// Mitsubishi GX Works2 project: TRANG TRAI BAN CU   PLC: FX3U/FX3UC

PROGRAM MAIN
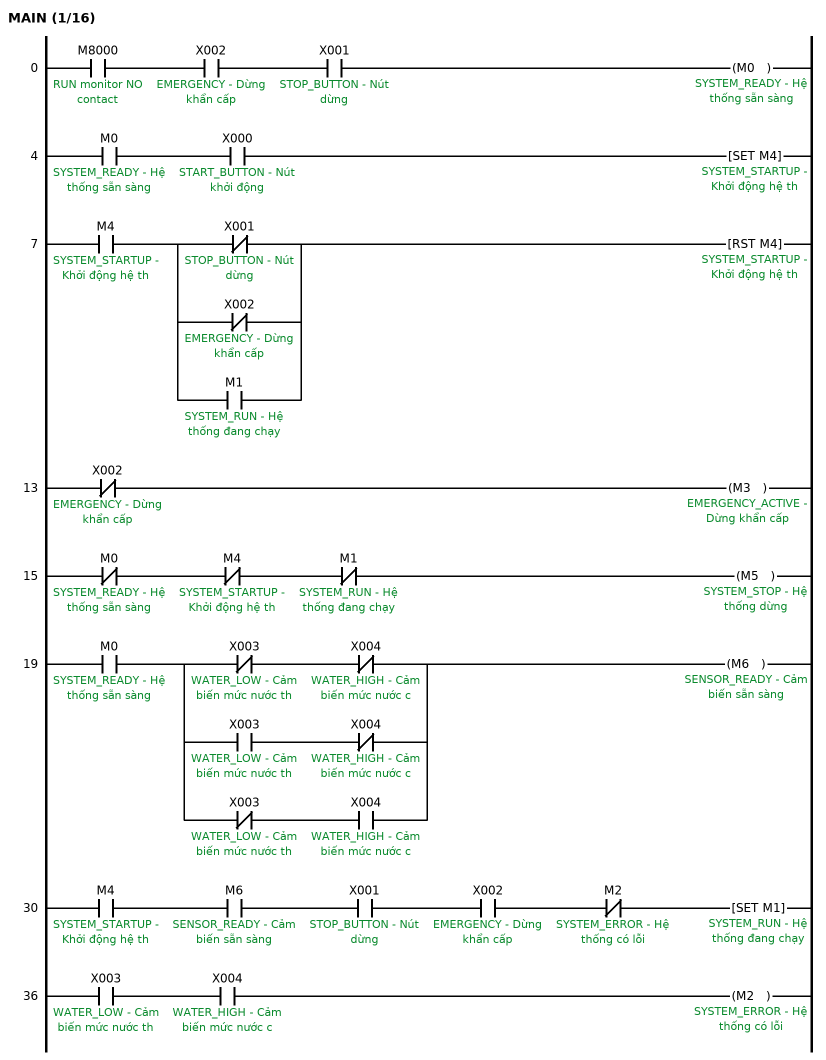
0     LD      M8000  ; RUN monitor NO contact
      AND     X002  ; EMERGENCY - Dừng khẩn cấp
      AND     X001  ; STOP_BUTTON - Nút dừng
      OUT     M0  ; SYSTEM_READY - Hệ thống sẵn sàng
4     LD      M0  ; SYSTEM_READY - Hệ thống sẵn sàng
      AND     X000  ; START_BUTTON - Nút khởi động
      SET     M4  ; SYSTEM_STARTUP - Khởi động hệ th
7     LD      M4  ; SYSTEM_STARTUP - Khởi động hệ th
      LDI     X001  ; STOP_BUTTON - Nút dừng
      ORI     X002  ; EMERGENCY - Dừng khẩn cấp
      OR      M1  ; SYSTEM_RUN - Hệ thống đang chạy
      ANB
      RST     M4  ; SYSTEM_STARTUP - Khởi động hệ th
13    LDI     X002  ; EMERGENCY - Dừng khẩn cấp
      OUT     M3  ; EMERGENCY_ACTIVE - Dừng khẩn cấp
15    LDI     M0  ; SYSTEM_READY - Hệ thống sẵn sàng
      ANI     M4  ; SYSTEM_STARTUP - Khởi động hệ th
      ANI     M1  ; SYSTEM_RUN - Hệ thống đang chạy
      OUT     M5  ; SYSTEM_STOP - Hệ thống dừng
19    LD      M0  ; SYSTEM_READY - Hệ thống sẵn sàng
      LDI     X003  ; WATER_LOW - Cảm biến mức nước th
      ANI     X004  ; WATER_HIGH - Cảm biến mức nước c
      LD      X003  ; WATER_LOW - Cảm biến mức nước th
      ANI     X004  ; WATER_HIGH - Cảm biến mức nước c
      ORB
      LDI     X003  ; WATER_LOW - Cảm biến mức nước th
      AND     X004  ; WATER_HIGH - Cảm biến mức nước c
      ORB
      ANB
      OUT     M6  ; SENSOR_READY - Cảm biến sẵn sàng
30    LD      M4  ; SYSTEM_STARTUP - Khởi động hệ th
      AND     M6  ; SENSOR_READY - Cảm biến sẵn sàng
      AND     X001  ; STOP_BUTTON - Nút dừng
      AND     X002  ; EMERGENCY - Dừng khẩn cấp
      ANI     M2  ; SYSTEM_ERROR - Hệ thống có lỗi
      SET     M1  ; SYSTEM_RUN - Hệ thống đang chạy
36    LD      X003  ; WATER_LOW - Cảm biến mức nước th
      AND     X004  ; WATER_HIGH - Cảm biến mức nước c
      OUT     M2  ; SYSTEM_ERROR - Hệ thống có lỗi
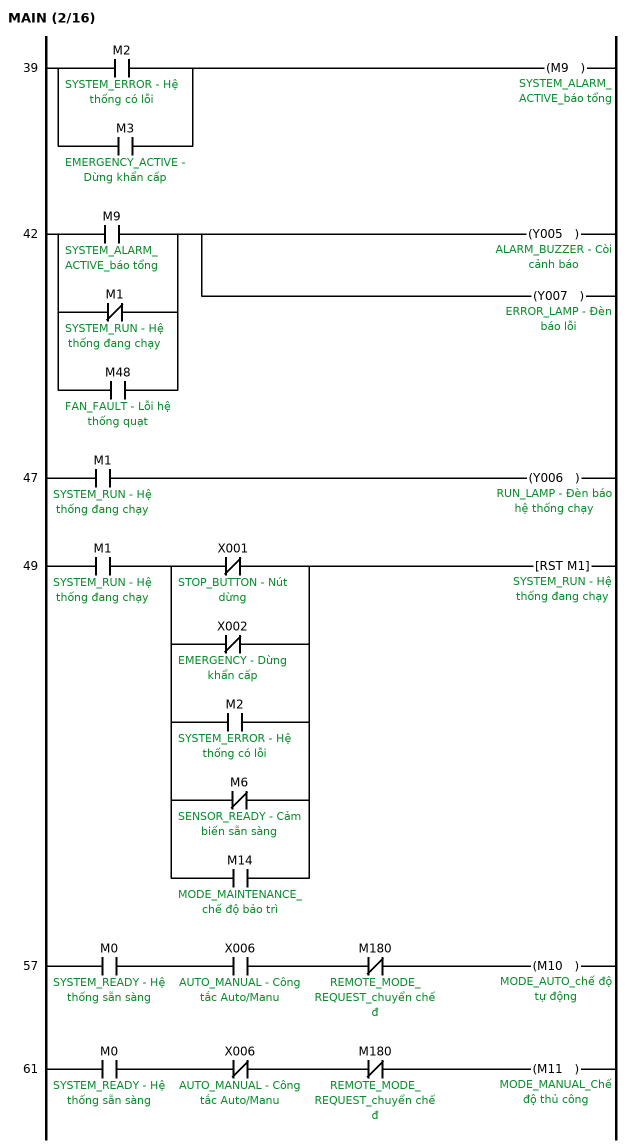
39    LD      M2  ; SYSTEM_ERROR - Hệ thống có lỗi
      OR      M3  ; EMERGENCY_ACTIVE - Dừng khẩn cấp
      OUT     M9  ; SYSTEM_ALARM_ACTIVE_báo tổng
42    LD      M9  ; SYSTEM_ALARM_ACTIVE_báo tổng
      ORI     M1  ; SYSTEM_RUN - Hệ thống đang chạy
      OR      M48  ; FAN_FAULT - Lỗi hệ thống quạt
      OUT     Y005  ; ALARM_BUZZER - Còi cảnh báo
      OUT     Y007  ; ERROR_LAMP - Đèn báo lỗi
47    LD      M1  ; SYSTEM_RUN - Hệ thống đang chạy
      OUT     Y006  ; RUN_LAMP - Đèn báo hệ thống chạy
49    LD      M1  ; SYSTEM_RUN - Hệ thống đang chạy
      LDI     X001  ; STOP_BUTTON - Nút dừng
      ORI     X002  ; EMERGENCY - Dừng khẩn cấp
      OR      M2  ; SYSTEM_ERROR - Hệ thống có lỗi
      ORI     M6  ; SENSOR_READY - Cảm biến sẵn sàng
      OR      M14  ; MODE_MAINTENANCE_chế độ bảo trì
      ANB
      RST     M1  ; SYSTEM_RUN - Hệ thống đang chạy
57    LD      M0  ; SYSTEM_READY - Hệ thống sẵn sàng
      AND     X006  ; AUTO_MANUAL - Công tắc Auto/Manu
      ANI     M180  ; REMOTE_MODE_REQUEST_chuyển chế đ
      OUT     M10  ; MODE_AUTO_chế độ tự động
61    LD      M0  ; SYSTEM_READY - Hệ thống sẵn sàng
      ANI     X006  ; AUTO_MANUAL - Công tắc Auto/Manu
      ANI     M180  ; REMOTE_MODE_REQUEST_chuyển chế đ
      OUT     M11  ; MODE_MANUAL_Chế độ thủ công
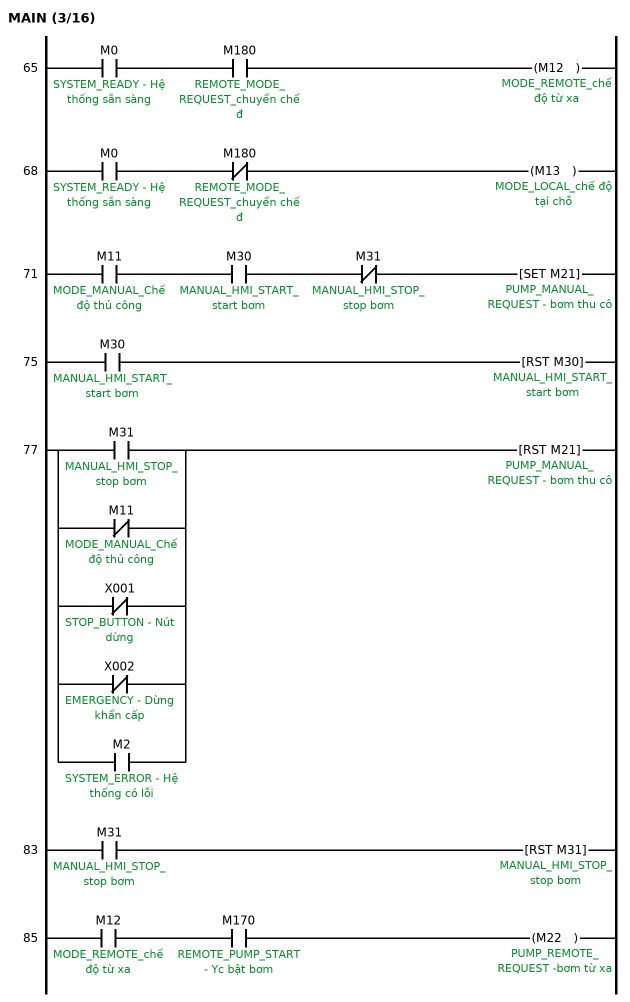
65    LD      M0  ; SYSTEM_READY - Hệ thống sẵn sàng
      AND     M180  ; REMOTE_MODE_REQUEST_chuyển chế đ
      OUT     M12  ; MODE_REMOTE_chế độ từ xa
68    LD      M0  ; SYSTEM_READY - Hệ thống sẵn sàng
      ANI     M180  ; REMOTE_MODE_REQUEST_chuyển chế đ
      OUT     M13  ; MODE_LOCAL_chế độ tại chỗ
71    LD      M11  ; MODE_MANUAL_Chế độ thủ công
      AND     M30  ; MANUAL_HMI_START_start bơm
      ANI     M31  ; MANUAL_HMI_STOP_stop bơm
      SET     M21  ; PUMP_MANUAL_REQUEST - bơm thu cô
75    LD      M30  ; MANUAL_HMI_START_start bơm
      RST     M30  ; MANUAL_HMI_START_start bơm
77    LD      M31  ; MANUAL_HMI_STOP_stop bơm
      ORI     M11  ; MODE_MANUAL_Chế độ thủ công
      ORI     X001  ; STOP_BUTTON - Nút dừng
      ORI     X002  ; EMERGENCY - Dừng khẩn cấp
      OR      M2  ; SYSTEM_ERROR - Hệ thống có lỗi
      RST     M21  ; PUMP_MANUAL_REQUEST - bơm thu cô
83    LD      M31  ; MANUAL_HMI_STOP_stop bơm
      RST     M31  ; MANUAL_HMI_STOP_stop bơm
85    LD      M12  ; MODE_REMOTE_chế độ từ xa
      AND     M170  ; REMOTE_PUMP_START - Yc bật bơm
      OUT     M22  ; PUMP_REMOTE_REQUEST -bơm từ xa
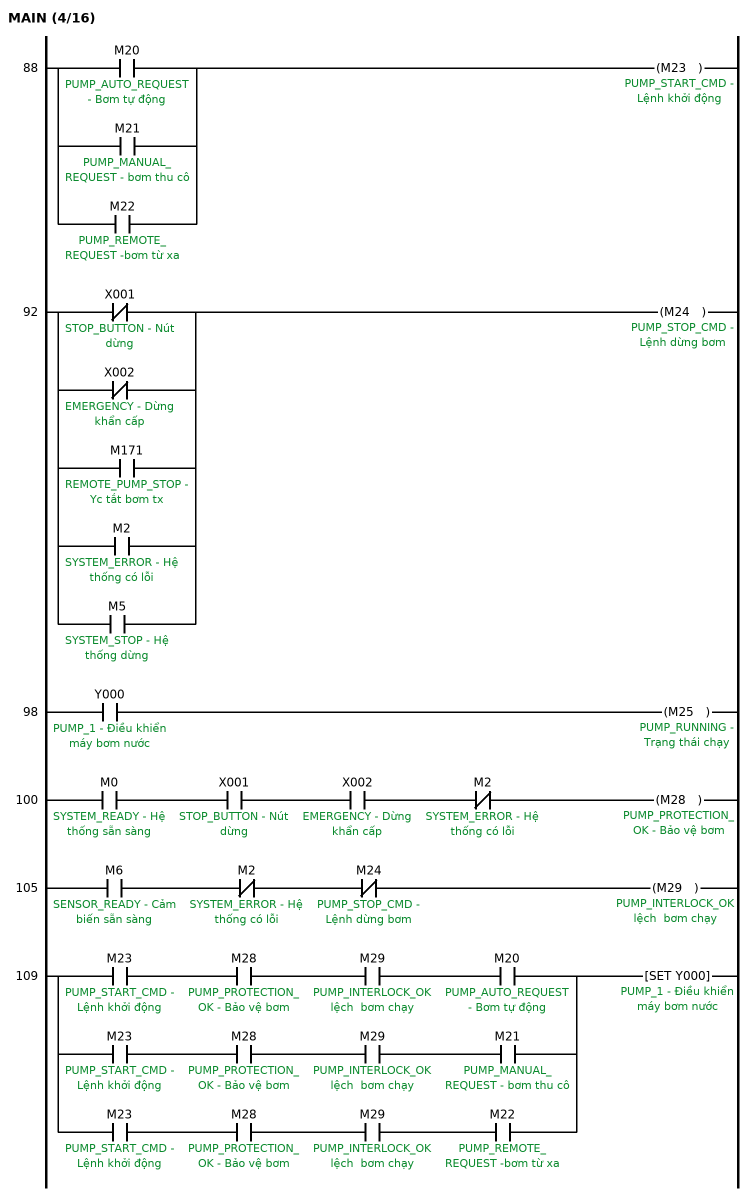
88    LD      M20  ; PUMP_AUTO_REQUEST - Bơm tự động
      OR      M21  ; PUMP_MANUAL_REQUEST - bơm thu cô
      OR      M22  ; PUMP_REMOTE_REQUEST -bơm từ xa
      OUT     M23  ; PUMP_START_CMD - Lệnh khởi động
92    LDI     X001  ; STOP_BUTTON - Nút dừng
      ORI     X002  ; EMERGENCY - Dừng khẩn cấp
      OR      M171  ; REMOTE_PUMP_STOP - Yc tắt bơm tx
      OR      M2  ; SYSTEM_ERROR - Hệ thống có lỗi
      OR      M5  ; SYSTEM_STOP - Hệ thống dừng
      OUT     M24  ; PUMP_STOP_CMD - Lệnh dừng bơm
98    LD      Y000  ; PUMP_1 - Điều khiển máy bơm nước
      OUT     M25  ; PUMP_RUNNING - Trạng thái chạy
100   LD      M0  ; SYSTEM_READY - Hệ thống sẵn sàng
      AND     X001  ; STOP_BUTTON - Nút dừng
      AND     X002  ; EMERGENCY - Dừng khẩn cấp
      ANI     M2  ; SYSTEM_ERROR - Hệ thống có lỗi
      OUT     M28  ; PUMP_PROTECTION_OK - Bảo vệ bơm
105   LD      M6  ; SENSOR_READY - Cảm biến sẵn sàng
      ANI     M2  ; SYSTEM_ERROR - Hệ thống có lỗi
      ANI     M24  ; PUMP_STOP_CMD - Lệnh dừng bơm
      OUT     M29  ; PUMP_INTERLOCK_OK lệch  bơm chạy
109   LD      M23  ; PUMP_START_CMD - Lệnh khởi động
      AND     M28  ; PUMP_PROTECTION_OK - Bảo vệ bơm
      AND     M29  ; PUMP_INTERLOCK_OK lệch  bơm chạy
      AND     M20  ; PUMP_AUTO_REQUEST - Bơm tự động
      LD      M23  ; PUMP_START_CMD - Lệnh khởi động
      AND     M28  ; PUMP_PROTECTION_OK - Bảo vệ bơm
      AND     M29  ; PUMP_INTERLOCK_OK lệch  bơm chạy
      AND     M21  ; PUMP_MANUAL_REQUEST - bơm thu cô
      ORB
      LD      M23  ; PUMP_START_CMD - Lệnh khởi động
      AND     M28  ; PUMP_PROTECTION_OK - Bảo vệ bơm
      AND     M29  ; PUMP_INTERLOCK_OK lệch  bơm chạy
      AND     M22  ; PUMP_REMOTE_REQUEST -bơm từ xa
      ORB
      SET     Y000  ; PUMP_1 - Điều khiển máy bơm nước
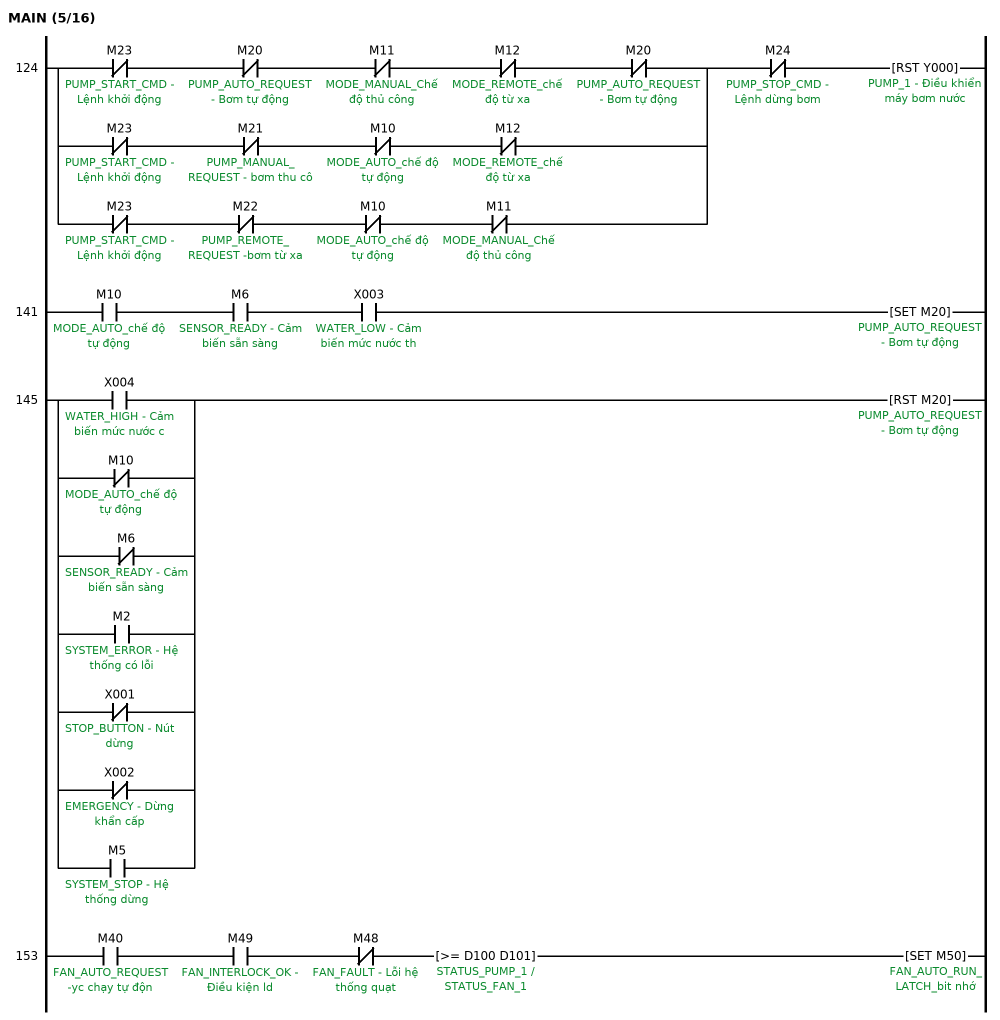
124   LDI     M23  ; PUMP_START_CMD - Lệnh khởi động
      ANI     M20  ; PUMP_AUTO_REQUEST - Bơm tự động
      ANI     M11  ; MODE_MANUAL_Chế độ thủ công
      ANI     M12  ; MODE_REMOTE_chế độ từ xa
      ANI     M20  ; PUMP_AUTO_REQUEST - Bơm tự động
      LDI     M23  ; PUMP_START_CMD - Lệnh khởi động
      ANI     M21  ; PUMP_MANUAL_REQUEST - bơm thu cô
      ANI     M10  ; MODE_AUTO_chế độ tự động
      ANI     M12  ; MODE_REMOTE_chế độ từ xa
      ORB
      LDI     M23  ; PUMP_START_CMD - Lệnh khởi động
      ANI     M22  ; PUMP_REMOTE_REQUEST -bơm từ xa
      ANI     M10  ; MODE_AUTO_chế độ tự động
      ANI     M11  ; MODE_MANUAL_Chế độ thủ công
      ORB
      ANI     M24  ; PUMP_STOP_CMD - Lệnh dừng bơm
      RST     Y000  ; PUMP_1 - Điều khiển máy bơm nước
141   LD      M10  ; MODE_AUTO_chế độ tự động
      AND     M6  ; SENSOR_READY - Cảm biến sẵn sàng
      AND     X003  ; WATER_LOW - Cảm biến mức nước th
      SET     M20  ; PUMP_AUTO_REQUEST - Bơm tự động
145   LD      X004  ; WATER_HIGH - Cảm biến mức nước c
      ORI     M10  ; MODE_AUTO_chế độ tự động
      ORI     M6  ; SENSOR_READY - Cảm biến sẵn sàng
      OR      M2  ; SYSTEM_ERROR - Hệ thống có lỗi
      ORI     X001  ; STOP_BUTTON - Nút dừng
      ORI     X002  ; EMERGENCY - Dừng khẩn cấp
      OR      M5  ; SYSTEM_STOP - Hệ thống dừng
      RST     M20  ; PUMP_AUTO_REQUEST - Bơm tự động
153   LD      M40  ; FAN_AUTO_REQUEST -yc chạy tự độn
      AND     M49  ; FAN_INTERLOCK_OK - Điều kiện ld
      ANI     M48  ; FAN_FAULT - Lỗi hệ thống quạt
      AND>=   D100 D101  ; STATUS_PUMP_1 / STATUS_FAN_1
      SET     M50  ; FAN_AUTO_RUN_LATCH_bit nhớ
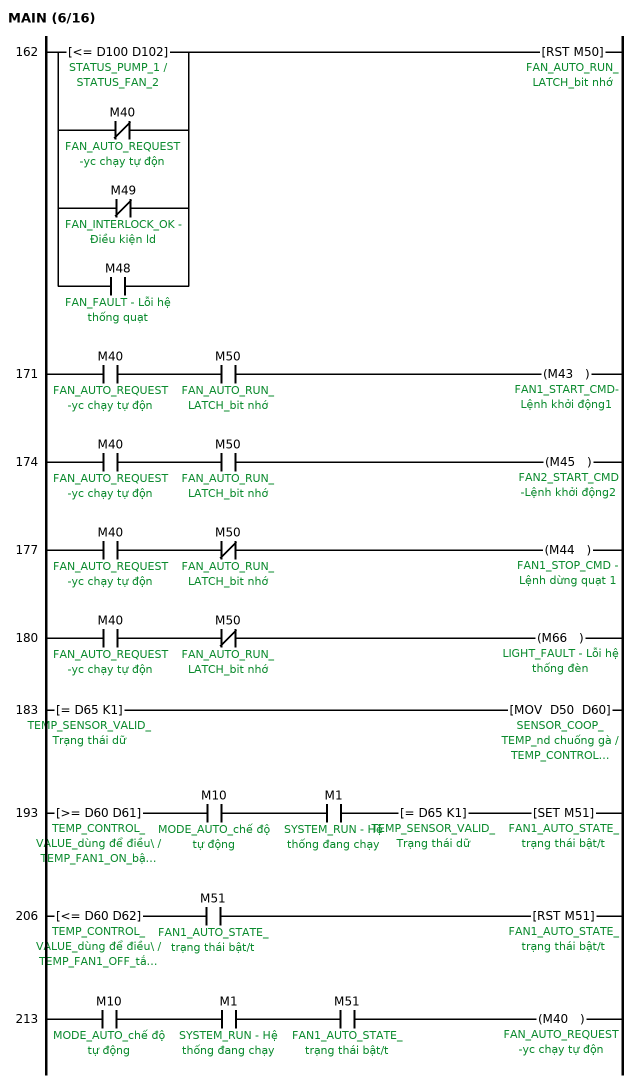
162   LD<=    D100 D102  ; STATUS_PUMP_1 / STATUS_FAN_2
      ORI     M40  ; FAN_AUTO_REQUEST -yc chạy tự độn
      ORI     M49  ; FAN_INTERLOCK_OK - Điều kiện ld
      OR      M48  ; FAN_FAULT - Lỗi hệ thống quạt
      RST     M50  ; FAN_AUTO_RUN_LATCH_bit nhớ
171   LD      M40  ; FAN_AUTO_REQUEST -yc chạy tự độn
      AND     M50  ; FAN_AUTO_RUN_LATCH_bit nhớ
      OUT     M43  ; FAN1_START_CMD-Lệnh khởi động1
174   LD      M40  ; FAN_AUTO_REQUEST -yc chạy tự độn
      AND     M50  ; FAN_AUTO_RUN_LATCH_bit nhớ
      OUT     M45  ; FAN2_START_CMD -Lệnh khởi động2
177   LD      M40  ; FAN_AUTO_REQUEST -yc chạy tự độn
      ANI     M50  ; FAN_AUTO_RUN_LATCH_bit nhớ
      OUT     M44  ; FAN1_STOP_CMD - Lệnh dừng quạt 1
180   LD      M40  ; FAN_AUTO_REQUEST -yc chạy tự độn
      ANI     M50  ; FAN_AUTO_RUN_LATCH_bit nhớ
      OUT     M66  ; LIGHT_FAULT - Lỗi hệ thống đèn
183   LD=     D65 K1  ; TEMP_SENSOR_VALID_Trạng thái dữ
      MOV     D50 D60  ; SENSOR_COOP_TEMP_nd chuống gà / TEMP_CONTROL_VALUE_dùng để điều\
193   LD>=    D60 D61  ; TEMP_CONTROL_VALUE_dùng để điều\ / TEMP_FAN1_ON_bật quạt 1
      AND     M10  ; MODE_AUTO_chế độ tự động
      AND     M1  ; SYSTEM_RUN - Hệ thống đang chạy
      AND=    D65 K1  ; TEMP_SENSOR_VALID_Trạng thái dữ
      SET     M51  ; FAN1_AUTO_STATE_trạng thái bật/t
206   LD<=    D60 D62  ; TEMP_CONTROL_VALUE_dùng để điều\ / TEMP_FAN1_OFF_tắt quạt 1
      AND     M51  ; FAN1_AUTO_STATE_trạng thái bật/t
      RST     M51  ; FAN1_AUTO_STATE_trạng thái bật/t
213   LD      M10  ; MODE_AUTO_chế độ tự động
      AND     M1  ; SYSTEM_RUN - Hệ thống đang chạy
      AND     M51  ; FAN1_AUTO_STATE_trạng thái bật/t
      OUT     M40  ; FAN_AUTO_REQUEST -yc chạy tự độn
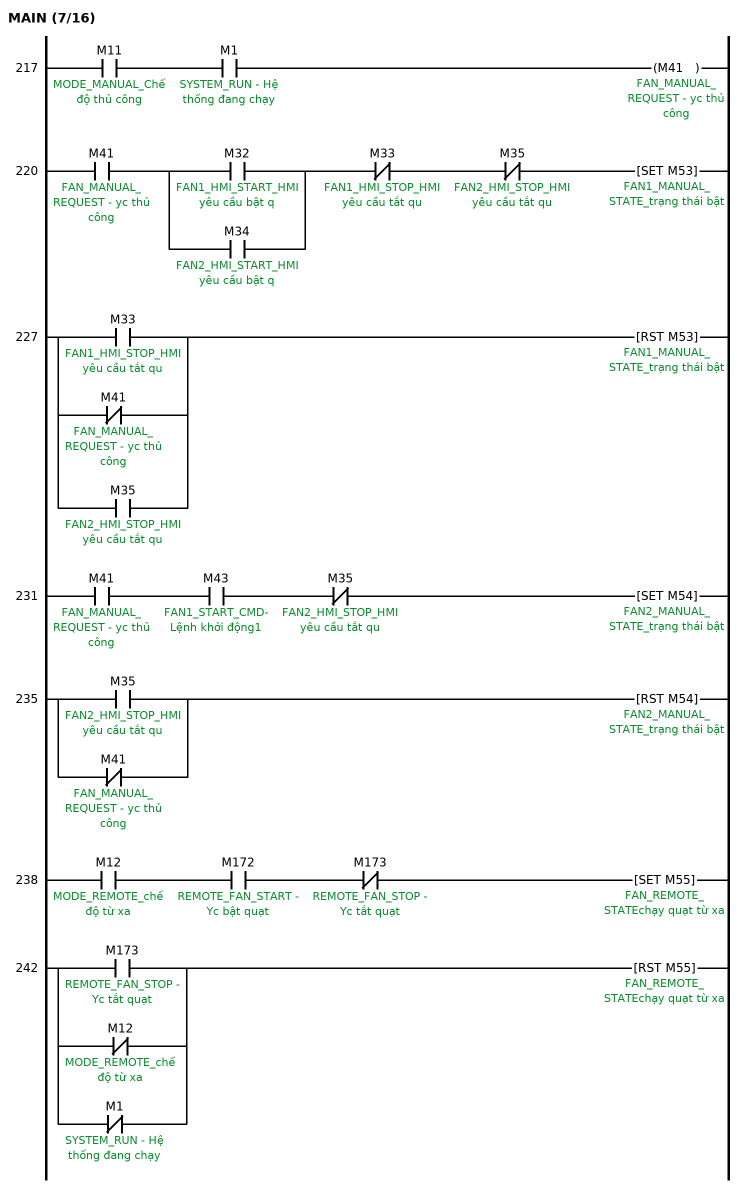
217   LD      M11  ; MODE_MANUAL_Chế độ thủ công
      AND     M1  ; SYSTEM_RUN - Hệ thống đang chạy
      OUT     M41  ; FAN_MANUAL_REQUEST - yc thủ công
220   LD      M41  ; FAN_MANUAL_REQUEST - yc thủ công
      LD      M32  ; FAN1_HMI_START_HMI yêu cầu bật q
      OR      M34  ; FAN2_HMI_START_HMI yêu cầu bật q
      ANB
      ANI     M33  ; FAN1_HMI_STOP_HMI yêu cầu tắt qu
      ANI     M35  ; FAN2_HMI_STOP_HMI yêu cầu tắt qu
      SET     M53  ; FAN1_MANUAL_STATE_trạng thái bật
227   LD      M33  ; FAN1_HMI_STOP_HMI yêu cầu tắt qu
      ORI     M41  ; FAN_MANUAL_REQUEST - yc thủ công
      OR      M35  ; FAN2_HMI_STOP_HMI yêu cầu tắt qu
      RST     M53  ; FAN1_MANUAL_STATE_trạng thái bật
231   LD      M41  ; FAN_MANUAL_REQUEST - yc thủ công
      AND     M43  ; FAN1_START_CMD-Lệnh khởi động1
      ANI     M35  ; FAN2_HMI_STOP_HMI yêu cầu tắt qu
      SET     M54  ; FAN2_MANUAL_STATE_trạng thái bật
235   LD      M35  ; FAN2_HMI_STOP_HMI yêu cầu tắt qu
      ORI     M41  ; FAN_MANUAL_REQUEST - yc thủ công
      RST     M54  ; FAN2_MANUAL_STATE_trạng thái bật
238   LD      M12  ; MODE_REMOTE_chế độ từ xa
      AND     M172  ; REMOTE_FAN_START - Yc bật quạt
      ANI     M173  ; REMOTE_FAN_STOP - Yc tắt quạt
      SET     M55  ; FAN_REMOTE_STATEchạy quạt từ xa
242   LD      M173  ; REMOTE_FAN_STOP - Yc tắt quạt
      ORI     M12  ; MODE_REMOTE_chế độ từ xa
      ORI     M1  ; SYSTEM_RUN - Hệ thống đang chạy
      RST     M55  ; FAN_REMOTE_STATEchạy quạt từ xa
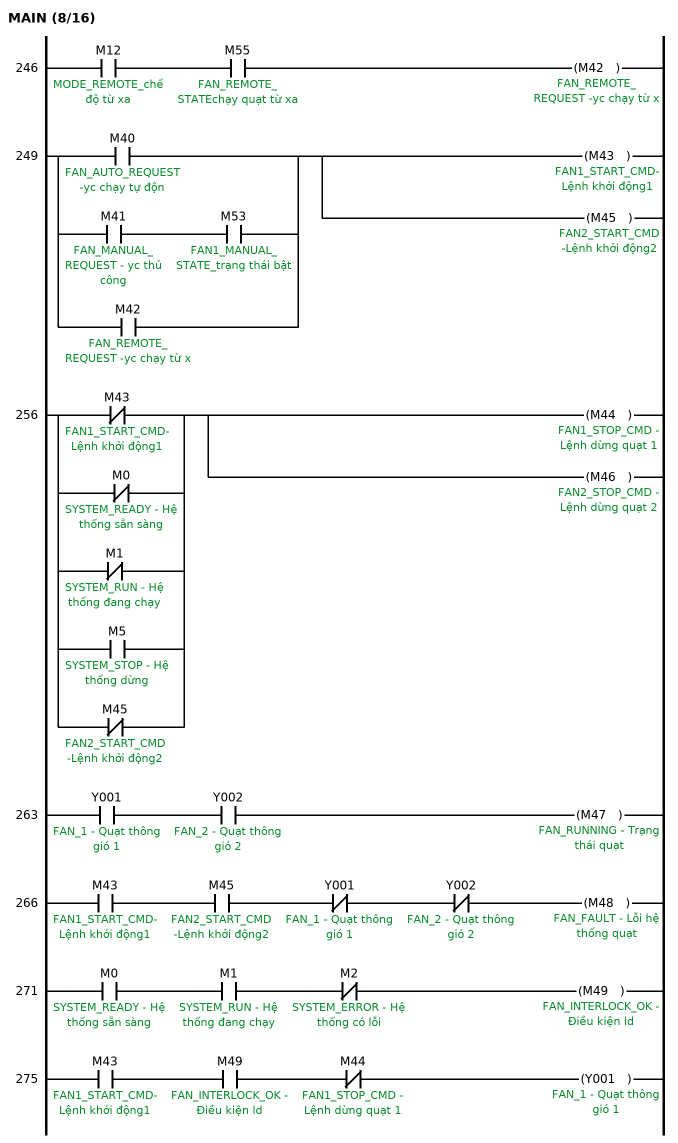
246   LD      M12  ; MODE_REMOTE_chế độ từ xa
      AND     M55  ; FAN_REMOTE_STATEchạy quạt từ xa
      OUT     M42  ; FAN_REMOTE_REQUEST -yc chạy từ x
249   LD      M40  ; FAN_AUTO_REQUEST -yc chạy tự độn
      LD      M41  ; FAN_MANUAL_REQUEST - yc thủ công
      AND     M53  ; FAN1_MANUAL_STATE_trạng thái bật
      ORB
      OR      M42  ; FAN_REMOTE_REQUEST -yc chạy từ x
      OUT     M43  ; FAN1_START_CMD-Lệnh khởi động1
      OUT     M45  ; FAN2_START_CMD -Lệnh khởi động2
256   LDI     M43  ; FAN1_START_CMD-Lệnh khởi động1
      ORI     M0  ; SYSTEM_READY - Hệ thống sẵn sàng
      ORI     M1  ; SYSTEM_RUN - Hệ thống đang chạy
      OR      M5  ; SYSTEM_STOP - Hệ thống dừng
      ORI     M45  ; FAN2_START_CMD -Lệnh khởi động2
      OUT     M44  ; FAN1_STOP_CMD - Lệnh dừng quạt 1
      OUT     M46  ; FAN2_STOP_CMD - Lệnh dừng quạt 2
263   LD      Y001  ; FAN_1 - Quạt thông gió 1
      AND     Y002  ; FAN_2 - Quạt thông gió 2
      OUT     M47  ; FAN_RUNNING - Trạng thái quạt
266   LD      M43  ; FAN1_START_CMD-Lệnh khởi động1
      AND     M45  ; FAN2_START_CMD -Lệnh khởi động2
      ANI     Y001  ; FAN_1 - Quạt thông gió 1
      ANI     Y002  ; FAN_2 - Quạt thông gió 2
      OUT     M48  ; FAN_FAULT - Lỗi hệ thống quạt
271   LD      M0  ; SYSTEM_READY - Hệ thống sẵn sàng
      AND     M1  ; SYSTEM_RUN - Hệ thống đang chạy
      ANI     M2  ; SYSTEM_ERROR - Hệ thống có lỗi
      OUT     M49  ; FAN_INTERLOCK_OK - Điều kiện ld
275   LD      M43  ; FAN1_START_CMD-Lệnh khởi động1
      AND     M49  ; FAN_INTERLOCK_OK - Điều kiện ld
      ANI     M44  ; FAN1_STOP_CMD - Lệnh dừng quạt 1
      OUT     Y001  ; FAN_1 - Quạt thông gió 1
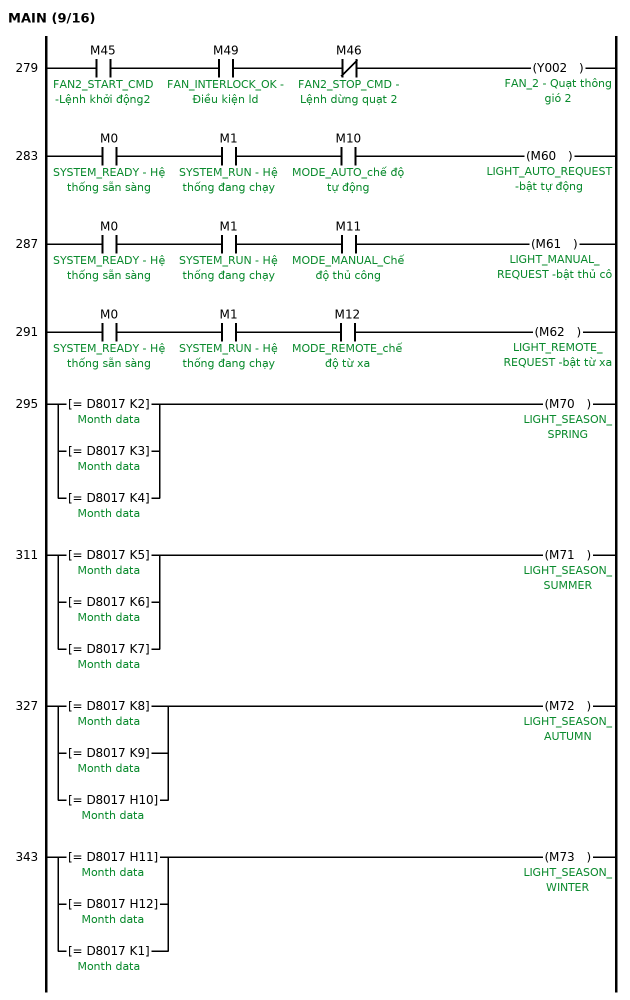
279   LD      M45  ; FAN2_START_CMD -Lệnh khởi động2
      AND     M49  ; FAN_INTERLOCK_OK - Điều kiện ld
      ANI     M46  ; FAN2_STOP_CMD - Lệnh dừng quạt 2
      OUT     Y002  ; FAN_2 - Quạt thông gió 2
283   LD      M0  ; SYSTEM_READY - Hệ thống sẵn sàng
      AND     M1  ; SYSTEM_RUN - Hệ thống đang chạy
      AND     M10  ; MODE_AUTO_chế độ tự động
      OUT     M60  ; LIGHT_AUTO_REQUEST -bật tự động
287   LD      M0  ; SYSTEM_READY - Hệ thống sẵn sàng
      AND     M1  ; SYSTEM_RUN - Hệ thống đang chạy
      AND     M11  ; MODE_MANUAL_Chế độ thủ công
      OUT     M61  ; LIGHT_MANUAL_REQUEST -bật thủ cô
291   LD      M0  ; SYSTEM_READY - Hệ thống sẵn sàng
      AND     M1  ; SYSTEM_RUN - Hệ thống đang chạy
      AND     M12  ; MODE_REMOTE_chế độ từ xa
      OUT     M62  ; LIGHT_REMOTE_REQUEST -bật từ xa
295   LD=     D8017 K2  ; Month data
      OR=     D8017 K3  ; Month data
      OR=     D8017 K4  ; Month data
      OUT     M70  ; LIGHT_SEASON_SPRING
311   LD=     D8017 K5  ; Month data
      OR=     D8017 K6  ; Month data
      OR=     D8017 K7  ; Month data
      OUT     M71  ; LIGHT_SEASON_SUMMER
327   LD=     D8017 K8  ; Month data
      OR=     D8017 K9  ; Month data
      OR=     D8017 H10  ; Month data
      OUT     M72  ; LIGHT_SEASON_AUTUMN
343   LD=     D8017 H11  ; Month data
      OR=     D8017 H12  ; Month data
      OR=     D8017 K1  ; Month data
      OUT     M73  ; LIGHT_SEASON_WINTER
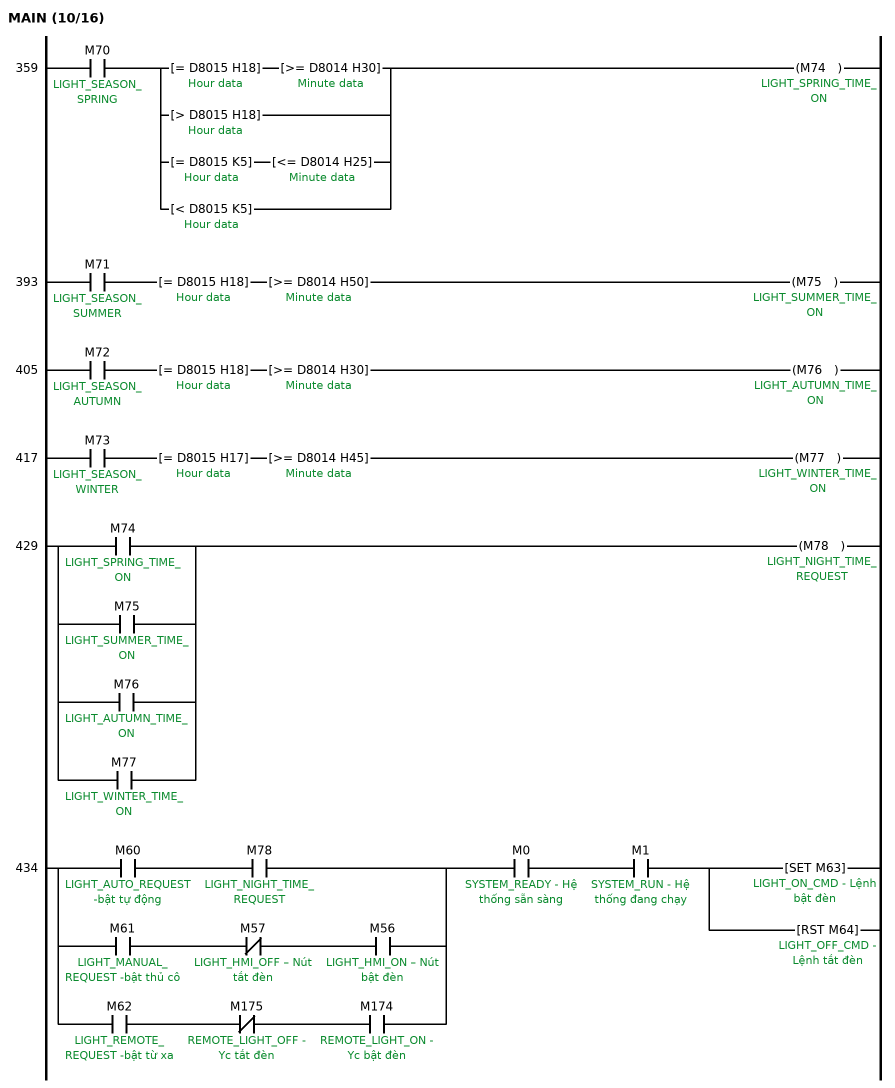
359   LD      M70  ; LIGHT_SEASON_SPRING
      LD=     D8015 H18  ; Hour data
      AND>=   D8014 H30  ; Minute data
      OR>     D8015 H18  ; Hour data
      LD=     D8015 K5  ; Hour data
      AND<=   D8014 H25  ; Minute data
      ORB
      OR<     D8015 K5  ; Hour data
      ANB
      OUT     M74  ; LIGHT_SPRING_TIME_ON
393   LD      M71  ; LIGHT_SEASON_SUMMER
      AND=    D8015 H18  ; Hour data
      AND>=   D8014 H50  ; Minute data
      OUT     M75  ; LIGHT_SUMMER_TIME_ON
405   LD      M72  ; LIGHT_SEASON_AUTUMN
      AND=    D8015 H18  ; Hour data
      AND>=   D8014 H30  ; Minute data
      OUT     M76  ; LIGHT_AUTUMN_TIME_ON
417   LD      M73  ; LIGHT_SEASON_WINTER
      AND=    D8015 H17  ; Hour data
      AND>=   D8014 H45  ; Minute data
      OUT     M77  ; LIGHT_WINTER_TIME_ON
429   LD      M74  ; LIGHT_SPRING_TIME_ON
      OR      M75  ; LIGHT_SUMMER_TIME_ON
      OR      M76  ; LIGHT_AUTUMN_TIME_ON
      OR      M77  ; LIGHT_WINTER_TIME_ON
      OUT     M78  ; LIGHT_NIGHT_TIME_REQUEST
434   LD      M60  ; LIGHT_AUTO_REQUEST -bật tự động
      AND     M78  ; LIGHT_NIGHT_TIME_REQUEST
      LD      M61  ; LIGHT_MANUAL_REQUEST -bật thủ cô
      ANI     M57  ; LIGHT_HMI_OFF – Nút tắt đèn
      AND     M56  ; LIGHT_HMI_ON – Nút bật đèn
      ORB
      LD      M62  ; LIGHT_REMOTE_REQUEST -bật từ xa
      ANI     M175  ; REMOTE_LIGHT_OFF - Yc tắt đèn
      AND     M174  ; REMOTE_LIGHT_ON - Yc bật đèn
      ORB
      AND     M0  ; SYSTEM_READY - Hệ thống sẵn sàng
      AND     M1  ; SYSTEM_RUN - Hệ thống đang chạy
      SET     M63  ; LIGHT_ON_CMD - Lệnh bật đèn
      RST     M64  ; LIGHT_OFF_CMD - Lệnh tắt đèn
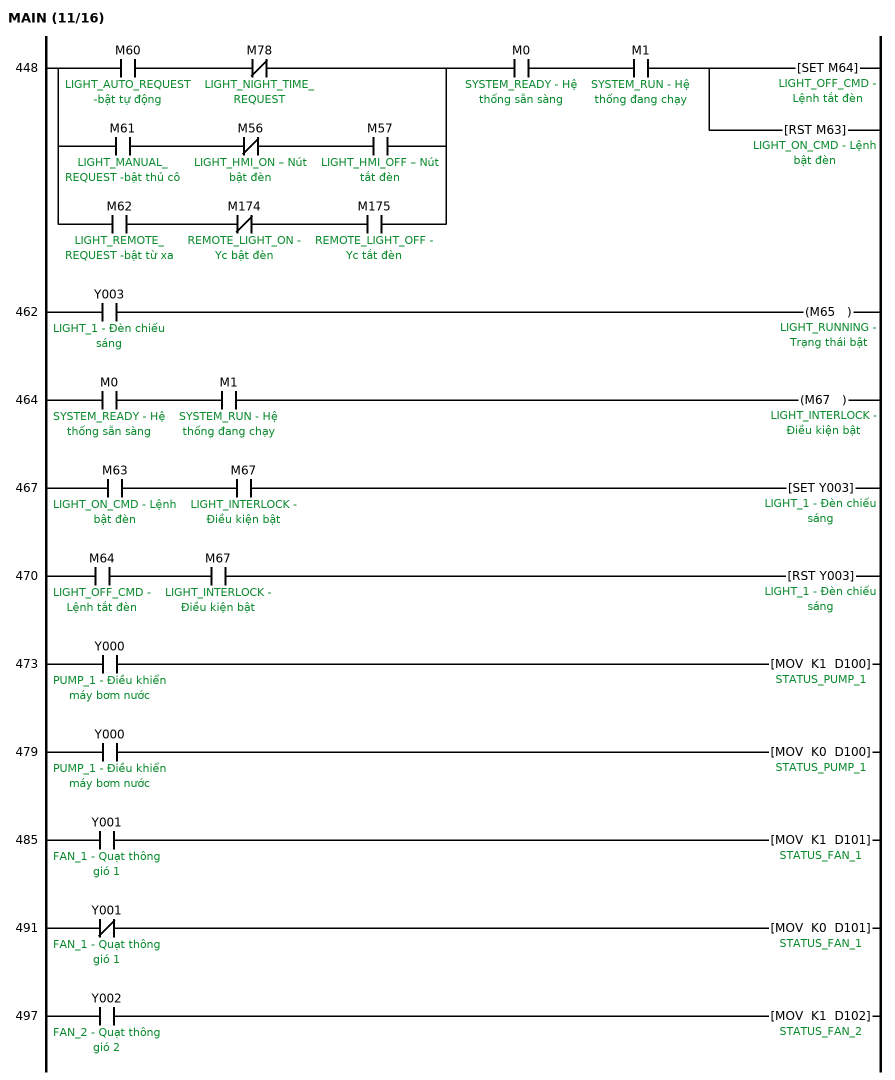
448   LD      M60  ; LIGHT_AUTO_REQUEST -bật tự động
      ANI     M78  ; LIGHT_NIGHT_TIME_REQUEST
      LD      M61  ; LIGHT_MANUAL_REQUEST -bật thủ cô
      ANI     M56  ; LIGHT_HMI_ON – Nút bật đèn
      AND     M57  ; LIGHT_HMI_OFF – Nút tắt đèn
      ORB
      LD      M62  ; LIGHT_REMOTE_REQUEST -bật từ xa
      ANI     M174  ; REMOTE_LIGHT_ON - Yc bật đèn
      AND     M175  ; REMOTE_LIGHT_OFF - Yc tắt đèn
      ORB
      AND     M0  ; SYSTEM_READY - Hệ thống sẵn sàng
      AND     M1  ; SYSTEM_RUN - Hệ thống đang chạy
      SET     M64  ; LIGHT_OFF_CMD - Lệnh tắt đèn
      RST     M63  ; LIGHT_ON_CMD - Lệnh bật đèn
462   LD      Y003  ; LIGHT_1 - Đèn chiếu sáng
      OUT     M65  ; LIGHT_RUNNING - Trạng thái bật
464   LD      M0  ; SYSTEM_READY - Hệ thống sẵn sàng
      AND     M1  ; SYSTEM_RUN - Hệ thống đang chạy
      OUT     M67  ; LIGHT_INTERLOCK - Điều kiện bật
467   LD      M63  ; LIGHT_ON_CMD - Lệnh bật đèn
      AND     M67  ; LIGHT_INTERLOCK - Điều kiện bật
      SET     Y003  ; LIGHT_1 - Đèn chiếu sáng
470   LD      M64  ; LIGHT_OFF_CMD - Lệnh tắt đèn
      AND     M67  ; LIGHT_INTERLOCK - Điều kiện bật
      RST     Y003  ; LIGHT_1 - Đèn chiếu sáng
473   LD      Y000  ; PUMP_1 - Điều khiển máy bơm nước
      MOV     K1 D100
479   LD      Y000  ; PUMP_1 - Điều khiển máy bơm nước
      MOV     K0 D100
485   LD      Y001  ; FAN_1 - Quạt thông gió 1
      MOV     K1 D101
491   LDI     Y001  ; FAN_1 - Quạt thông gió 1
      MOV     K0 D101
497   LD      Y002  ; FAN_2 - Quạt thông gió 2
      MOV     K1 D102
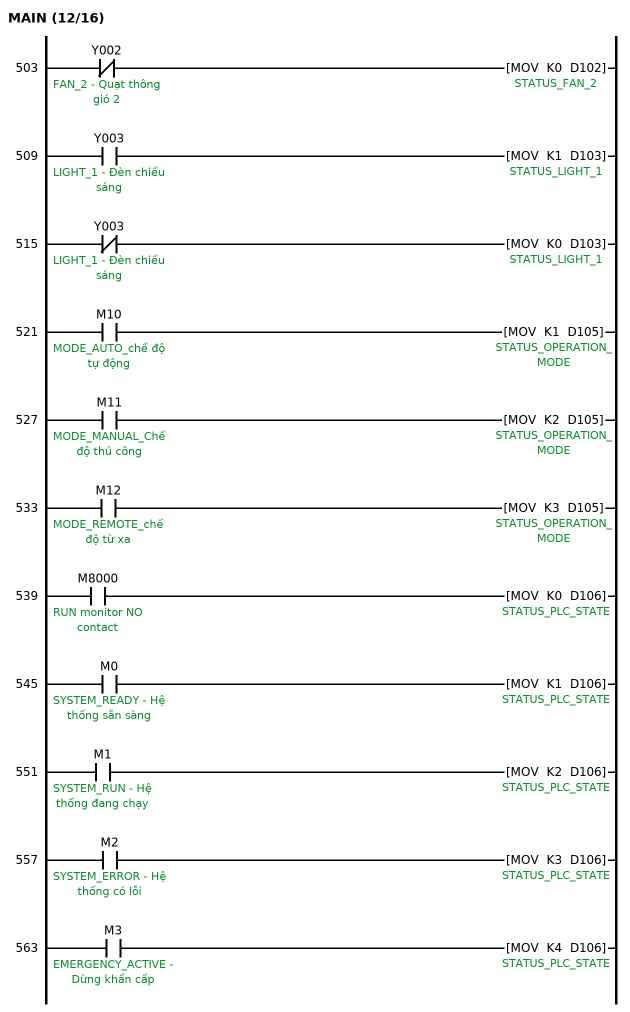
503   LDI     Y002  ; FAN_2 - Quạt thông gió 2
      MOV     K0 D102
509   LD      Y003  ; LIGHT_1 - Đèn chiếu sáng
      MOV     K1 D103  ; STATUS_LIGHT_1
515   LDI     Y003  ; LIGHT_1 - Đèn chiếu sáng
      MOV     K0 D103
521   LD      M10  ; MODE_AUTO_chế độ tự động
      MOV     K1 D105  ; STATUS_OPERATION_MODE
527   LD      M11  ; MODE_MANUAL_Chế độ thủ công
      MOV     K2 D105
533   LD      M12  ; MODE_REMOTE_chế độ từ xa
      MOV     K3 D105
539   LD      M8000  ; RUN monitor NO contact
      MOV     K0 D106  ; STATUS_PLC_STATE
545   LD      M0  ; SYSTEM_READY - Hệ thống sẵn sàng
      MOV     K1 D106
551   LD      M1  ; SYSTEM_RUN - Hệ thống đang chạy
      MOV     K2 D106
557   LD      M2  ; SYSTEM_ERROR - Hệ thống có lỗi
      MOV     K3 D106
563   LD      M3  ; EMERGENCY_ACTIVE - Dừng khẩn cấp
      MOV     K4 D106
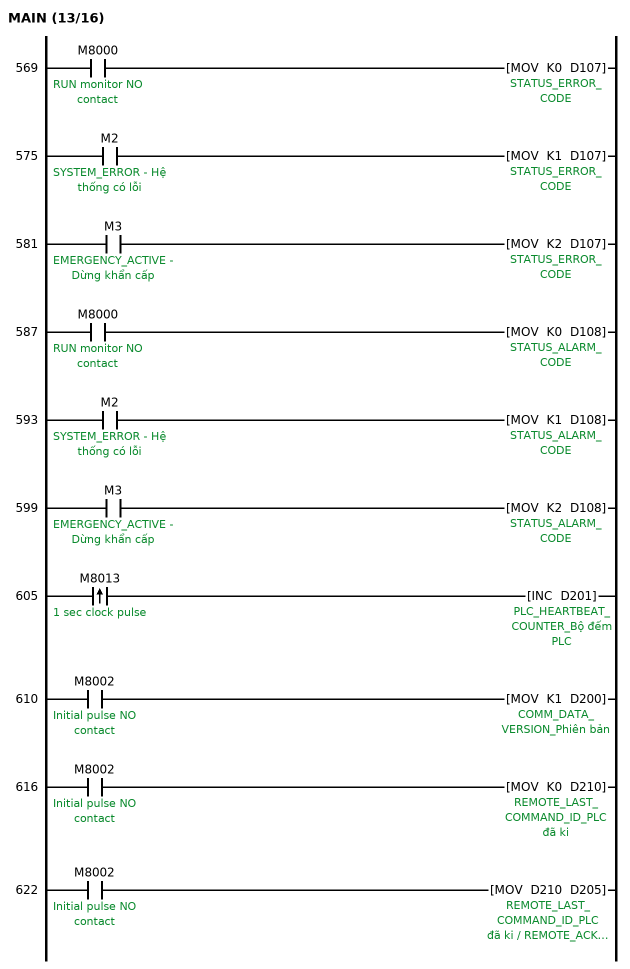
569   LD      M8000  ; RUN monitor NO contact
      MOV     K0 D107  ; STATUS_ERROR_CODE
575   LD      M2  ; SYSTEM_ERROR - Hệ thống có lỗi
      MOV     K1 D107
581   LD      M3  ; EMERGENCY_ACTIVE - Dừng khẩn cấp
      MOV     K2 D107
587   LD      M8000  ; RUN monitor NO contact
      MOV     K0 D108  ; STATUS_ALARM_CODE
593   LD      M2  ; SYSTEM_ERROR - Hệ thống có lỗi
      MOV     K1 D108
599   LD      M3  ; EMERGENCY_ACTIVE - Dừng khẩn cấp
      MOV     K2 D108
605   LDP     M8013  ; 1 sec clock pulse
      INC     D201  ; PLC_HEARTBEAT_COUNTER_Bộ đếm PLC
610   LD      M8002  ; Initial pulse NO contact
      MOV     K1 D200  ; COMM_DATA_VERSION_Phiên bản
616   LD      M8002  ; Initial pulse NO contact
      MOV     K0 D210  ; REMOTE_LAST_COMMAND_ID_PLC đã ki
622   LD      M8002  ; Initial pulse NO contact
      MOV     D210 D205  ; REMOTE_ACK_COMMAND_ID_PLC đã nhậ
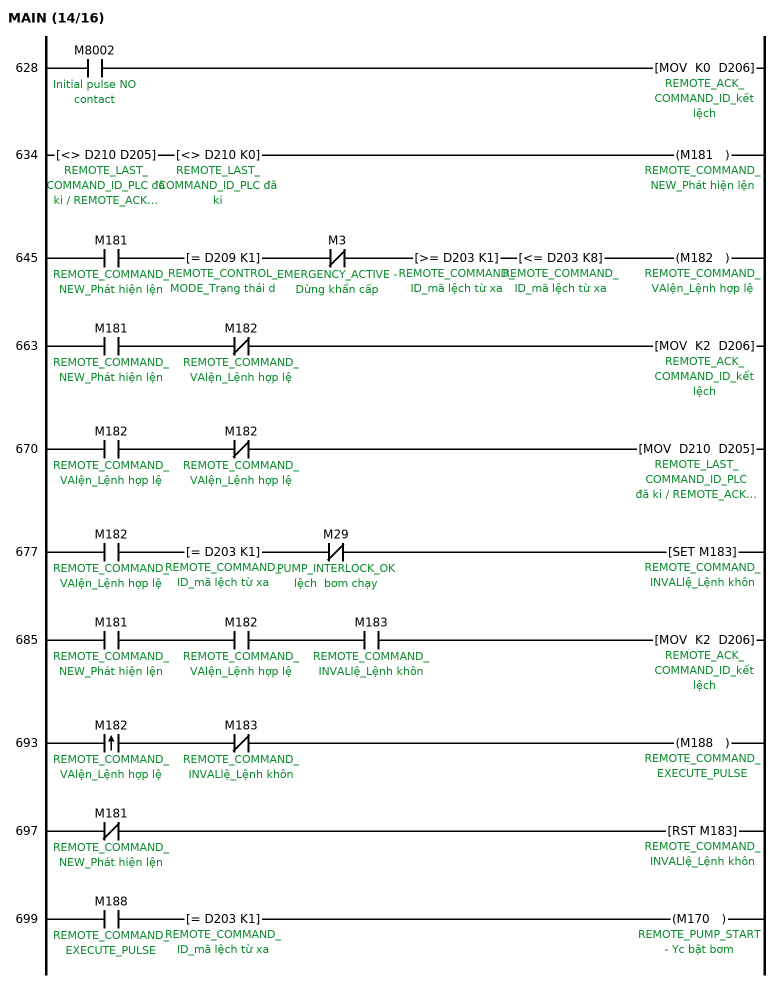
628   LD      M8002  ; Initial pulse NO contact
      MOV     K0 D206  ; REMOTE_ACK_COMMAND_ID_kết lệch
634   LD<>    D210 D205  ; REMOTE_LAST_COMMAND_ID_PLC đã ki / REMOTE_ACK_COMMAND_ID_PLC đã nhậ
      AND<>   D210 K0  ; REMOTE_LAST_COMMAND_ID_PLC đã ki
      OUT     M181  ; REMOTE_COMMAND_NEW_Phát hiện lện
645   LD      M181  ; REMOTE_COMMAND_NEW_Phát hiện lện
      AND=    D209 K1  ; REMOTE_CONTROL_MODE_Trạng thái d
      ANI     M3  ; EMERGENCY_ACTIVE - Dừng khẩn cấp
      AND>=   D203 K1  ; REMOTE_COMMAND_ID_mã lệch từ xa
      AND<=   D203 K8  ; REMOTE_COMMAND_ID_mã lệch từ xa
      OUT     M182  ; REMOTE_COMMAND_VAlện_Lệnh hợp lệ
663   LD      M181  ; REMOTE_COMMAND_NEW_Phát hiện lện
      ANI     M182  ; REMOTE_COMMAND_VAlện_Lệnh hợp lệ
      MOV     K2 D206
670   LD      M182  ; REMOTE_COMMAND_VAlện_Lệnh hợp lệ
      ANI     M182  ; REMOTE_COMMAND_VAlện_Lệnh hợp lệ
      MOV     D210 D205
677   LD      M182  ; REMOTE_COMMAND_VAlện_Lệnh hợp lệ
      AND=    D203 K1  ; REMOTE_COMMAND_ID_mã lệch từ xa
      ANI     M29  ; PUMP_INTERLOCK_OK lệch  bơm chạy
      SET     M183  ; REMOTE_COMMAND_INVALlệ_Lệnh khôn
685   LD      M181  ; REMOTE_COMMAND_NEW_Phát hiện lện
      AND     M182  ; REMOTE_COMMAND_VAlện_Lệnh hợp lệ
      AND     M183  ; REMOTE_COMMAND_INVALlệ_Lệnh khôn
      MOV     K2 D206
693   LDP     M182  ; REMOTE_COMMAND_VAlện_Lệnh hợp lệ
      ANI     M183  ; REMOTE_COMMAND_INVALlệ_Lệnh khôn
      OUT     M188  ; REMOTE_COMMAND_EXECUTE_PULSE
697   LDI     M181  ; REMOTE_COMMAND_NEW_Phát hiện lện
      RST     M183  ; REMOTE_COMMAND_INVALlệ_Lệnh khôn
699   LD      M188  ; REMOTE_COMMAND_EXECUTE_PULSE
      AND=    D203 K1  ; REMOTE_COMMAND_ID_mã lệch từ xa
      OUT     M170  ; REMOTE_PUMP_START - Yc bật bơm
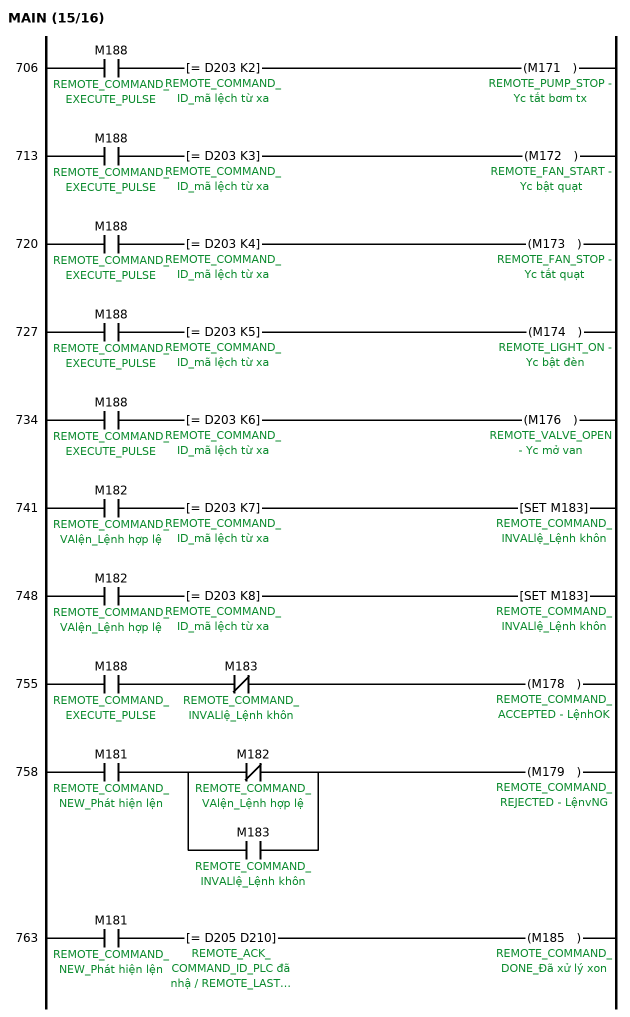
706   LD      M188  ; REMOTE_COMMAND_EXECUTE_PULSE
      AND=    D203 K2  ; REMOTE_COMMAND_ID_mã lệch từ xa
      OUT     M171  ; REMOTE_PUMP_STOP - Yc tắt bơm tx
713   LD      M188  ; REMOTE_COMMAND_EXECUTE_PULSE
      AND=    D203 K3  ; REMOTE_COMMAND_ID_mã lệch từ xa
      OUT     M172  ; REMOTE_FAN_START - Yc bật quạt
720   LD      M188  ; REMOTE_COMMAND_EXECUTE_PULSE
      AND=    D203 K4  ; REMOTE_COMMAND_ID_mã lệch từ xa
      OUT     M173  ; REMOTE_FAN_STOP - Yc tắt quạt
727   LD      M188  ; REMOTE_COMMAND_EXECUTE_PULSE
      AND=    D203 K5  ; REMOTE_COMMAND_ID_mã lệch từ xa
      OUT     M174  ; REMOTE_LIGHT_ON - Yc bật đèn
734   LD      M188  ; REMOTE_COMMAND_EXECUTE_PULSE
      AND=    D203 K6  ; REMOTE_COMMAND_ID_mã lệch từ xa
      OUT     M176  ; REMOTE_VALVE_OPEN - Yc mở van
741   LD      M182  ; REMOTE_COMMAND_VAlện_Lệnh hợp lệ
      AND=    D203 K7  ; REMOTE_COMMAND_ID_mã lệch từ xa
      SET     M183  ; REMOTE_COMMAND_INVALlệ_Lệnh khôn
748   LD      M182  ; REMOTE_COMMAND_VAlện_Lệnh hợp lệ
      AND=    D203 K8  ; REMOTE_COMMAND_ID_mã lệch từ xa
      SET     M183  ; REMOTE_COMMAND_INVALlệ_Lệnh khôn
755   LD      M188  ; REMOTE_COMMAND_EXECUTE_PULSE
      ANI     M183  ; REMOTE_COMMAND_INVALlệ_Lệnh khôn
      OUT     M178  ; REMOTE_COMMAND_ACCEPTED - LệnhOK
758   LD      M181  ; REMOTE_COMMAND_NEW_Phát hiện lện
      LDI     M182  ; REMOTE_COMMAND_VAlện_Lệnh hợp lệ
      OR      M183  ; REMOTE_COMMAND_INVALlệ_Lệnh khôn
      ANB
      OUT     M179  ; REMOTE_COMMAND_REJECTED - LệnvNG
763   LD      M181  ; REMOTE_COMMAND_NEW_Phát hiện lện
      AND=    D205 D210  ; REMOTE_ACK_COMMAND_ID_PLC đã nhậ / REMOTE_LAST_COMMAND_ID_PLC đã ki
      OUT     M185  ; REMOTE_COMMAND_DONE_Đã xử lý xon
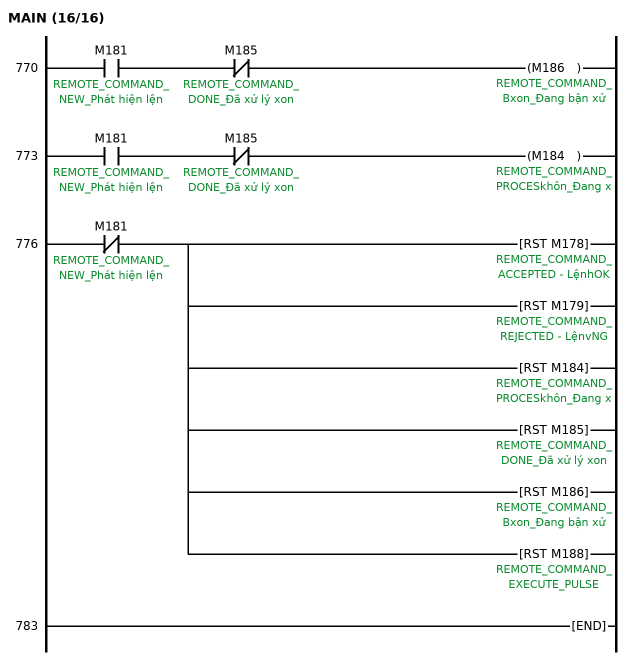
770   LD      M181  ; REMOTE_COMMAND_NEW_Phát hiện lện
      ANI     M185  ; REMOTE_COMMAND_DONE_Đã xử lý xon
      OUT     M186  ; REMOTE_COMMAND_Bxon_Đang bận xử
773   LD      M181  ; REMOTE_COMMAND_NEW_Phát hiện lện
      ANI     M185  ; REMOTE_COMMAND_DONE_Đã xử lý xon
      OUT     M184  ; REMOTE_COMMAND_PROCESkhôn_Đang x
776   LDI     M181  ; REMOTE_COMMAND_NEW_Phát hiện lện
      RST     M178  ; REMOTE_COMMAND_ACCEPTED - LệnhOK
      RST     M179  ; REMOTE_COMMAND_REJECTED - LệnvNG
      RST     M184  ; REMOTE_COMMAND_PROCESkhôn_Đang x
      RST     M185  ; REMOTE_COMMAND_DONE_Đã xử lý xon
      RST     M186  ; REMOTE_COMMAND_Bxon_Đang bận xử
      RST     M188  ; REMOTE_COMMAND_EXECUTE_PULSE
783   END
END_PROGRAM

// device comments not shown above
X005  ; DOOR_SENSOR - Cảm biến cửa
Y004  ; VALVE_1 - Van cấp nước
M7  ; AUTO_ENABLE - Cho phép chế độ tự
M8  ; MANUAL_ENABLE - Cho phép chế độ
M15  ; MODE_INITIALIZING_Trạng thái HT
M26  ; PUMP_FAULT - Lỗi máy bơm
M27  ; PUMP_TIMEOUT - Bơm chạy quá
M52  ; FAN2_AUTO_STATE_trạng thái bật/t
M80  ; VALVE_AUTO_REQUEST_mở tự động
M81  ; VALVE_MANUAL_REQUEST -mở thủ côn
M82  ; VALVE_REMOTE_REQUEST -mở từ xa
M83  ; VALVE_OPEN_CMD - Lệnh mở van
M84  ; VALVE_CLOSE_CMD - Lệnh đóng van
M85  ; VALVE_OPENING - Trạng thái mở
M86  ; VALVE_FAULT - Lỗi van cấp nước
M87  ; VALVE_INTERLOCK- Điều kiện mở
M88  ; WATER_SUPPLY_ACTIVE - Đang cấp n
M89  ; VALVE_TIMEOUT - Van hd quá giờ
M100  ; ALARM_TEMP_HIGH - Cảnh báo nhiệt
M101  ; ALARM_WATER_LOW - Cảnh báo mức t
M102  ; ALARM_PUMP_TIMEOUT_bơm quá giờ
M103  ; ALARM_FAN_FAULT - Cảnh báo quạt
M104  ; ALARM_SENSOR_FAULT -lỗi cảm biến
M105  ; ALARM_GATEWAY_OFFLINE -mất kết n
M106  ; ALARM_WATER_HIGH - nước quá cao
M107  ; ALARM_DOOR_OPEN - Cảnh báo cửa m
M108  ; ALARM_POWER_FAIL - mất nguồn
M109  ; ALARM_GENERAL - Cảnh báo tổng
M130  ; ERROR_TEMP_SENSOR - Lỗi cb nhiệt
M131  ; ERROR_HUMIDITY_SENSOR - Lỗi da
M132  ; ERROR_WATER_SENSOR - Lỗi cb mực
M133  ; ERROR_PUMP - Lỗi máy bơm
M134  ; ERROR_FAN - Lỗi quạt
M135  ; ERROR_VALVE - Lỗi van nước
M136  ; ERROR_GATEWAY - Lỗi Gateway
M137  ; ERROR_COMMUNICATION - Lỗi RS485
M138  ; ERROR_OVERLOAD - Lỗi quá tải thi
M139  ; ERROR_SYSTEM - Lỗi tổng hệ thống
M150  ; GATEWAY_ONLINE - Gateway kết nối
M151  ; GATEWAY_COMMAND_VALID - Lệnh OK
M152  ; GATEWAY_DATA_READY - Dữ liệu SS
M153  ; RS485_TX_REQUEST - gửi dữ liệu
M154  ; RS485_RX_COMPLETE - Nhận dữ liệu
M155  ; RS485_COMM_ERROR - Lỗi RS485
M156  ; PLC_HEARTBEAT - Xung kiểm traPLC
M157  ; GATEWAY_HEARTBEAT -kiểm tra gate
M158  ; COMM_TIMEOUT - Quá thời gian phả
M159  ; COMM_RECOVERY - Đã khôi phục kết
M177  ; REMOTE_VALVE_CLOSE - Yc đóng van
M187  ; REMOTE_COMMAND_RESET_Xóa trạng t
D0  ; SET_TEMP_FAN_ON_nd bật quạt
D1  ; SET_TEMP_FAN_OFF_nd tắt quạt
D2  ; SET_WATER_PUMP_ON_m bật bơm
D3  ; SET_WATER_PUMP_OFF_m tắt bơm
D4  ; SET_PUMP_MAX_TIME_tg bơm
D5  ; SET_ALARM_DELAY_thời gian trễ
D6  ; SET_TEMP_ALARM_HIGH_nhiệt độ cao
D7  ; SET_HUMIDITY_HIGH_độ âm cao
D8  ; SET_HUMIDITY_LOW_độ ẩm thấp
D9  ; SET_LIGHT_ON_TIME_bật đèn theo g
D10  ; SET_TEMP_ALARM_LOW_nhiệt độ thấ
D51  ; SENSOR_AIR_HUMIDITY_độ ẩm
D52  ; SENSOR_WATER_TEMP_nhiệt độ nước
D53  ; SENSOR_WATER_LEVEL_mực nước
D54  ; SENSOR_SOIL_HUMIDITY_độ ẩm đất
D55  ; SENSOR_LIGHT_VALUE_độ sáng
D56  ; SENSOR_CO2_VALUE_Nồng độ CO₂
D57  ; SENSOR_NH3_VALUE_Nồng độ NH₃
D58  ; SENSOR_TEMP_STATUS_trạng thái cb
D59  ; SENSOR_DATA_STATUS_trạng thái dl
D63  ; TEMP_FAN2_ON_bật quạt 2
D64  ; TEMP_FAN2_OFF_tắt quạt 2
D66  ; FAN_AUTO_DELAY_Thời gian trễ
D67  ; FAN_CONTROL_MODE_Chế độ điều khi
D68  ; FAN1_RUNTIME_Thời gian hoạt động
D69  ; FAN2_RUNTIME_Thời gian hoạt động
D104  ; STATUS_VALVE_1
D109  ; STATUS_SYSTEM_UPTIME
D202  ; GATEWAY_HEARTBEAT_COUNTER_gate
D204  ; REMOTE_COMMAND_VALUE_giá trị DK
D207  ; COMM_ERROR_CODE_Mã lỗi truyền th
D208  ; COMM_DATA_COUNTER_Bộ đếm dữ liệu
D300  ; STAT_PUMP_START_COUNT_số lần bơm
D301  ; STAT_PUMP_RUNTIME_MIN_hời gian b
D302  ; STAT_FAN_RUNTIME_MIN_tg quạt
D303  ; STAT_LIGHT_RUNTIME_MIN_tg bật đè
D304  ; STAT_VALVE_OPEN_COUNT_số lần mở
D305  ; STAT_ALARM_COUNT_số lần cảnh báo
D306  ; STAT_ERROR_COUNT_số lần lỗi
D307  ; STAT_GATEWAY_LOSS_COUNT_kết nối
D308  ; STAT_SENSOR_ERROR_COUNT_lỗi CB
D309  ; STAT_SYSTEM_RUNTIME_HOUR_giờ HD
